(*
SPDX-FileCopyrightText: © 2026 Oleksandr Tiutyk <trofimich@gmail.com>
SPDX-License-Identifier: MIT
License: https://opensource.org/license/mit
*)

(*!
<summary>Reports an error occurring during filesystem operations.</summary>
<description>
Reports caller-detected filesystem failures using the GeneralException lifetime and throw rules. Message is
borrowed read-only during the call; errorCode stores the native/ADS error identifier. Dynamic instances and
clones belong to DynamicMemoryManager until task cleanup. Plain __NEW does not transfer ownership to the task
manager.
</description>
*)

{attribute 'enable_dynamic_creation'}
{attribute 'no_explicit_call' := 'do not call this function block directly'}
FUNCTION_BLOCK FileSystemException EXTENDS TOF_Core.GeneralException IMPLEMENTS IFileSystemException
VAR_STAT
	{attribute 'hide'} 
	_ClassName : STRING := __POUNAME();
END_VAR

(*!
<summary>Provides the concrete type name used in diagnostics.</summary>
<description>
Returns borrowed read-only metadata; keep the instance alive and do not modify the referenced string.
Reading does not allocate memory, initialize resources or transfer ownership.
</description>
*)
{attribute 'monitoring' := 'call'}
PROPERTY ClassName : REFERENCE TO STRING
GET
ClassName REF= _ClassName;
END_GET
END_PROPERTY

(*!
<summary>Creates a task-owned copy of this exception and its diagnostic payload.</summary>
<description>
Registers the newly constructed instance before copying payload, outside FB_init. Registration failure
releases the unregistered instance and raises a terminal error; copy failure leaves the registered instance
owned by the task manager for cleanup. Custom overrides must follow the same ownership sequence. The returned
reference is borrowed until task cleanup and must not be deleted by the caller.
</description>
*)
METHOD Clone : TOF_Core.IObject
VAR
	exceptionClone : POINTER TO FileSystemException;
END_VAR
exceptionClone := __NEW(FileSystemException);

IF exceptionClone = 0 THEN
	TOF_Core.DynamicMemoryManager.RaiseAllocationFailure();
END_IF

TOF_Core.DynamicMemoryManager.RegisterAutoDisposedObject(autoDisposedObject := exceptionClone^);

exceptionClone^.CopyGeneralFields(sourceException := THIS^);

Clone := exceptionClone^;
END_METHOD

(*!
<summary>Provides the library namespace used in diagnostics.</summary>
<description>Returns borrowed read-only namespace storage; do not modify the referenced string.</description>
*)
{attribute 'monitoring' := 'call'}
PROPERTY NamespaceName : REFERENCE TO STRING
GET
NamespaceName REF= CurrentNamespace.Name;
END_GET
END_PROPERTY

(*!
<summary>Reports the size of this concrete instance in bytes.</summary>
*)
{attribute 'monitoring' := 'call'}
PROPERTY SelfSize : ULINT
GET
SelfSize := XSIZEOF(THIS^);
END_GET
END_PROPERTY

(*!
<summary>Raises a filesystem exception with the supplied message and error code.</summary>
<description>
Borrows message read-only for this call and records the numeric error code. Formats diagnostic text without
heap allocation during message preparation; does not retain the input reference. The caller detects the
filesystem error; this method propagates it.
</description>
<param name="sourceNamespaceName">Namespace of the caller.</param>
<param name="sourceClassName">Class name of the caller.</param>
<param name="sourcePOUName">POU name of the caller.</param>
<param name="sourcePosition">Source position of the caller.</param>
<param name="message">Diagnostic explanation.</param>
<param name="errorCode">Native/ADS error code, or 0 if unassigned.</param>
*)
METHOD Throw
VAR_INPUT
	sourceNamespaceName : STRING;
	sourceClassName : STRING;
	sourcePOUName : STRING;
	sourcePosition : STRING;
END_VAR
VAR_IN_OUT CONSTANT
	message : TOF_Core.ERROR_MESSAGE;
END_VAR
VAR_INPUT
	errorCode : UDINT := 0;
END_VAR
InternalThrow(
	sourceNamespaceName := sourceNamespaceName,
	sourceClassName := sourceClassName,
	sourcePOUName := sourcePOUName,
	sourcePosition := sourcePosition,
	message := message,
	errorCode := errorCode,
	innerException := 0
);
END_METHOD

END_FUNCTION_BLOCK

(* stored: Version 1.1.0.1
   POU FileSystemException: Id {ae1bbb4c-25c9-4ede-b477-d4e2dbf3bbcb}, SpecialFunc None
   Property ClassName: Id {376ea995-58b5-4c78-90b1-69650a357d0d}
   Get Get: Id {80c7e1c5-bd06-4d91-a5f8-ba7a9104a58f}
   Method Clone: Id {e792337e-6253-4b91-87c8-846b83c3e742}
   Property NamespaceName: Id {e661210f-f8c8-4dcc-89b3-816483dc0fc7}
   Get Get: Id {5fc180fe-9746-4cb8-bd97-0a075e11695c}
   Property SelfSize: Id {bbfec0e7-f859-42a0-936a-da63ff5b72d3}
   Get Get: Id {11aae084-3af3-48d8-b045-b79955e6f600}
   Method Throw: Id {1f875777-9d21-4766-ab74-aa42509cccbd} *)
